{attribute 'qualified_only'}
{attribute 'strict'}
TYPE E_CIP_TankList :
(
	eT91_Sanitation :=0,
	eT92_Detergent,
	eT93_R_Water,
	eT94_Water
);
END_TYPE

(* stored: Version 1.1.0.1, ProductVersion 3.1.4024.12
   DUT E_CIP_TankList: Id {8b6fc95d-14e2-474d-95b3-abd3db69964a} *)
